(*
SPDX-FileCopyrightText: © 2026 Oleksandr Tiutyk <trofimich@gmail.com>
SPDX-License-Identifier: MIT
License: https://opensource.org/license/mit
*)

(*!
<summary>Mock leaf for lifecycle hooks, I/O phases, initialization/reset faults and event routing.</summary>
*)

FUNCTION_BLOCK MockLeafAutomationComponent EXTENDS TOF_Automation.InputOutputLeafAutomationComponent
VAR_INPUT
	//! <summary>Raises one output fault after the output call has been counted.</summary>
	ThrowOnNextOutput : BOOL;
	//! <summary>Raises one fault during input acquisition.</summary>
	ThrowOnNextInput : BOOL;
END_VAR
VAR_STAT
	{attribute 'hide'}
	_ClassName : STRING := __POUNAME();
END_VAR
VAR
	{attribute 'hide'}
	_InitializeCount : INT;
	{attribute 'hide'}
	_WorkingCount : INT;
	{attribute 'hide'}
	_ProcessInputCount : INT;
	{attribute 'hide'}
	_ProcessOutputCount : INT;
	{attribute 'hide'}
	_ResetCount : INT;
	{attribute 'hide'}
	_StopCount : INT;
	{attribute 'hide'}
	_EnableCount : INT;
	{attribute 'hide'}
	_DisableCount : INT;
	{attribute 'hide'}
	_EventReceivedCount : INT;
	{attribute 'hide'}
	_LastReceivedEventId : INT;
	{attribute 'hide'}
	_StopPropagationOnEvent : BOOL;
	{attribute 'hide'}
	_InitReturnValue : BOOL := TRUE;
	{attribute 'hide'}
	_FailOnWorking : BOOL;
	_ThrowOnInitializing : BOOL;
	_ThrowOnReset : BOOL;
	_RecoverCount : INT;
	_ThrowOnRecover : BOOL;
	_ThrowOnEnable : BOOL;
	_ThrowOnDisable : BOOL;
END_VAR

{attribute 'monitoring' := 'call'}
PROPERTY ClassName : REFERENCE TO STRING
GET
ClassName REF= _ClassName;
END_GET
END_PROPERTY

{attribute 'monitoring' := 'call'}
PROPERTY DisableCount : INT
GET
DisableCount := _DisableCount;
END_GET
END_PROPERTY

{attribute 'monitoring' := 'call'}
PROPERTY EnableCount : INT
GET
EnableCount := _EnableCount;
END_GET
END_PROPERTY

{attribute 'monitoring' := 'call'}
PROPERTY EventReceivedCount : INT
GET
EventReceivedCount := _EventReceivedCount;
END_GET
END_PROPERTY

{attribute 'monitoring' := 'call'}
PROPERTY FailOnWorking : BOOL
GET
FailOnWorking := _FailOnWorking;
END_GET
SET
_FailOnWorking := FailOnWorking;
END_SET
END_PROPERTY

METHOD FB_init : BOOL
VAR_INPUT
	bInitRetains : BOOL; // TRUE: the retain variables are initialized (reset warm / reset cold)
	bInCopyCode : BOOL;  // TRUE: the instance will be copied to the copy code afterward (online change)
	name : WSTRING;
	parent : TOF_Automation.IParentAutomationComponent;
END_VAR
END_METHOD

{attribute 'monitoring' := 'call'}
PROPERTY InitializeCount : INT
GET
InitializeCount := _InitializeCount;
END_GET
END_PROPERTY

{attribute 'monitoring' := 'call'}
PROPERTY InitReturnValue : BOOL
GET
InitReturnValue := _InitReturnValue;
END_GET
SET
_InitReturnValue := InitReturnValue;
END_SET
END_PROPERTY

{attribute 'monitoring' := 'call'}
PROPERTY LastReceivedEventId : INT
GET
LastReceivedEventId := _LastReceivedEventId;
END_GET
END_PROPERTY

{attribute 'monitoring' := 'call'}
PROPERTY NamespaceName : REFERENCE TO STRING
GET
NamespaceName REF= CurrentNamespace.Name;
END_GET
END_PROPERTY

(*!
<summary>Records the OnDisable call and optionally injects an exception.</summary>
*)
METHOD PROTECTED OnDisable
_DisableCount := _DisableCount + 1;

IF _ThrowOnDisable THEN
	TOF_Core.Exceptions.ThrowStandard(
		sourceNamespaceName := NamespaceName,
		sourceClassName := ClassName,
		sourcePOUName := __POUNAME(),
		sourcePosition := __POSITION(),
		message := "Injected OnDisable failure."
	);
END_IF
END_METHOD

(*!
<summary>Records the OnEnable call and optionally injects an exception.</summary>
*)
METHOD PROTECTED OnEnable
_EnableCount := _EnableCount + 1;

IF _ThrowOnEnable THEN
	TOF_Core.Exceptions.ThrowStandard(
		sourceNamespaceName := NamespaceName,
		sourceClassName := ClassName,
		sourcePOUName := __POUNAME(),
		sourcePosition := __POSITION(),
		message := "Injected OnEnable failure."
	);
END_IF
END_METHOD

METHOD OnEventReceived
VAR_INPUT
	event : TOF_Core.IEvent;
END_VAR
VAR_OUTPUT
	stopPropagation : BOOL;
END_VAR
VAR
	mockEv : POINTER TO MockAutomationEvent;
END_VAR
_EventReceivedCount := _EventReceivedCount + 1;

IF __QUERYPOINTER(event, mockEv) THEN
	_LastReceivedEventId := mockEv^.EventId;
END_IF

stopPropagation := _StopPropagationOnEvent;
END_METHOD

(*!
<summary>Records the OnInitializing call and optionally injects an exception.</summary>
<description>
The exception exercises production conversion into a copied component error; the hook does not own it.
</description>
*)
METHOD PROTECTED OnInitializing : BOOL
_InitializeCount := _InitializeCount + 1;

IF _ThrowOnInitializing THEN
	TOF_Core.Exceptions.ThrowStandard(
		sourceNamespaceName := NamespaceName,
		sourceClassName := ClassName,
		sourcePOUName := __POUNAME(),
		sourcePosition := __POSITION(),
		message := "Injected OnInitializing failure."
	);
END_IF

OnInitializing := _InitReturnValue;
END_METHOD

(*! <summary>Counts input calls and raises an armed input fault once.</summary> *)
METHOD PROTECTED OnProcessInput
_ProcessInputCount := _ProcessInputCount + 1;

IF ThrowOnNextInput THEN
	ThrowOnNextInput := FALSE;
	TOF_Core.Exceptions.ThrowStandard(
		sourceNamespaceName := NamespaceName,
		sourceClassName := ClassName,
		sourcePOUName := __POUNAME(),
		sourcePosition := __POSITION(),
		message := "Injected input failure"
	);
END_IF
END_METHOD

(*! <summary>Counts output calls and optionally injects a one-shot fault after the observed effect.</summary> *)
METHOD PROTECTED OnProcessOutput
_ProcessOutputCount := _ProcessOutputCount + 1;

IF ThrowOnNextOutput THEN
	ThrowOnNextOutput := FALSE;
	TOF_Core.Exceptions.ThrowStandard(
		sourceNamespaceName := NamespaceName,
		sourceClassName := ClassName,
		sourcePOUName := __POUNAME(),
		sourcePosition := __POSITION(),
		message := "Injected output failure"
	);
END_IF
END_METHOD

(*!
<summary>Records the OnRecover call and optionally injects an exception.</summary>
*)
METHOD PROTECTED OnRecover
_RecoverCount := _RecoverCount + 1;

IF _ThrowOnRecover THEN
	TOF_Core.Exceptions.ThrowStandard(
		sourceNamespaceName := NamespaceName,
		sourceClassName := ClassName,
		sourcePOUName := __POUNAME(),
		sourcePosition := __POSITION(),
		message := "Injected OnRecover failure."
	);
END_IF
END_METHOD

(*!
<summary>Records the OnReset call and optionally injects an exception.</summary>
<description>
The exception exercises production conversion into a copied component error; the hook does not own it.
</description>
*)
METHOD PROTECTED OnReset
_ResetCount := _ResetCount + 1;

IF _ThrowOnReset THEN
	TOF_Core.Exceptions.ThrowStandard(
		sourceNamespaceName := NamespaceName,
		sourceClassName := ClassName,
		sourcePOUName := __POUNAME(),
		sourcePosition := __POSITION(),
		message := "Injected OnReset failure."
	);
END_IF
END_METHOD

METHOD PROTECTED OnStopped
_StopCount := _StopCount + 1;
END_METHOD

METHOD PROTECTED OnWorking
_WorkingCount := _WorkingCount + 1;

IF _FailOnWorking THEN
	TOF_Core.Exceptions.ThrowStandard(
		sourceNamespaceName := NamespaceName,
		sourceClassName := ClassName,
		sourcePOUName := __POUNAME(),
		sourcePosition := __POSITION(),
		message := "Mock leaf failure on working"
	);
END_IF
END_METHOD

{attribute 'monitoring' := 'call'}
PROPERTY ProcessInputCount : INT
GET
ProcessInputCount := _ProcessInputCount;
END_GET
END_PROPERTY

{attribute 'monitoring' := 'call'}
PROPERTY ProcessOutputCount : INT
GET
ProcessOutputCount := _ProcessOutputCount;
END_GET
END_PROPERTY

{attribute 'monitoring' := 'call'}
PROPERTY ResetCount : INT
GET
ResetCount := _ResetCount;
END_GET
END_PROPERTY

{attribute 'monitoring' := 'call'}
PROPERTY SelfSize : ULINT
GET
SelfSize := XSIZEOF(THIS^);
END_GET
END_PROPERTY

{attribute 'monitoring' := 'call'}
PROPERTY StopCount : INT
GET
StopCount := _StopCount;
END_GET
END_PROPERTY

{attribute 'monitoring' := 'call'}
PROPERTY StopPropagationOnEvent : BOOL
GET
StopPropagationOnEvent := _StopPropagationOnEvent;
END_GET
SET
_StopPropagationOnEvent := StopPropagationOnEvent;
END_SET
END_PROPERTY

{attribute 'monitoring' := 'call'}
PROPERTY WorkingCount : INT
GET
WorkingCount := _WorkingCount;
END_GET
END_PROPERTY

(*!
<summary>Controls the initialization-hook failure injected by regression tests.</summary>
*)
{attribute 'monitoring' := 'call'}
PROPERTY ThrowOnInitializing : BOOL
GET
ThrowOnInitializing := _ThrowOnInitializing;
END_GET
SET
_ThrowOnInitializing := ThrowOnInitializing;
END_SET
END_PROPERTY

(*!
<summary>Controls the reset-hook failure injected by regression tests.</summary>
*)
{attribute 'monitoring' := 'call'}
PROPERTY ThrowOnReset : BOOL
GET
ThrowOnReset := _ThrowOnReset;
END_GET
SET
_ThrowOnReset := ThrowOnReset;
END_SET
END_PROPERTY

(*!
<summary>Gets the number of OnRecover calls recorded by this mock leaf.</summary>
*)
{attribute 'monitoring' := 'call'}
PROPERTY RecoverCount : INT
GET
RecoverCount := _RecoverCount;
END_GET
END_PROPERTY

(*!
<summary>Controls the disable-hook failure injected by regression tests.</summary>
*)
{attribute 'monitoring' := 'call'}
PROPERTY ThrowOnDisable : BOOL
GET
ThrowOnDisable := _ThrowOnDisable;
END_GET
SET
_ThrowOnDisable := ThrowOnDisable;
END_SET
END_PROPERTY

(*!
<summary>Controls the enable-hook failure injected by regression tests.</summary>
*)
{attribute 'monitoring' := 'call'}
PROPERTY ThrowOnEnable : BOOL
GET
ThrowOnEnable := _ThrowOnEnable;
END_GET
SET
_ThrowOnEnable := ThrowOnEnable;
END_SET
END_PROPERTY

(*!
<summary>Controls the recover-hook failure injected by regression tests.</summary>
*)
{attribute 'monitoring' := 'call'}
PROPERTY ThrowOnRecover : BOOL
GET
ThrowOnRecover := _ThrowOnRecover;
END_GET
SET
_ThrowOnRecover := ThrowOnRecover;
END_SET
END_PROPERTY

(*!
<summary>Exercises the inherited exception handler with a borrowed diagnostic in the fixture's current state.</summary>
<param name="exception">Task-local exception that remains live for the call.</param>
<param name="reaction">Runtime reaction to apply.</param>
*)
METHOD ApplyExceptionReaction
VAR_INPUT
	exception : TOF_Core.IException;
	reaction : TOF_Core.EXCEPTION_REACTION;
END_VAR
ProcessException(exception := exception, exceptionReaction := reaction, exceptionSourceHint := "Injected primary failure");
END_METHOD

END_FUNCTION_BLOCK

(* stored: Version 1.1.0.1, ProductVersion 3.1.4026.21
   POU MockLeafAutomationComponent: Id {9b7b3daa-f346-4584-a906-6da16219c11f}, SpecialFunc None
   Folder Methods to override: Id {612da229-f7d8-494f-8591-082c05072b3f}
   Folder Properties for tests: Id {ccac3e62-bc35-4f89-a40e-c876ffb73e34}
   Property ClassName: Id {d5c4d5ee-cde5-4df4-8cbd-46cced7d5454}
   Get Get: Id {5415ed35-e09f-4119-8198-c8575e6b1ab5}
   Property DisableCount: Id {bbaaaf6d-9d95-455d-b78d-b03325aec8ca}
   Get Get: Id {16fe8a7f-cfad-4055-9144-48f18add74a5}
   Property EnableCount: Id {8454a8af-ef78-4131-b582-201baa06e86e}
   Get Get: Id {489c43e4-5062-4c21-8691-e46ab060d4b5}
   Property EventReceivedCount: Id {803a68c5-6fea-4132-9ec0-3eab19c89d39}
   Get Get: Id {bd615afb-6d2f-41d6-88ec-30cdcef21a93}
   Property FailOnWorking: Id {4ac1dd38-5fe7-40fa-b603-9534ebe240bd}
   Get Get: Id {da42525c-79be-4472-94c1-fd35af010373}
   Set Set: Id {a2eba756-0bc3-4394-adfb-aa16c4171792}
   Method FB_init: Id {2ce54561-f6b4-4f38-b28c-e9e2d5ba5306}
   Property InitializeCount: Id {ff7ba116-c221-4cd9-9799-5b16792aeb45}
   Get Get: Id {018cb720-e3f7-4649-8b67-bed593899c5b}
   Property InitReturnValue: Id {69a85714-ee34-4f3d-80b7-d8d28b5786a9}
   Get Get: Id {c7fd5de5-7d8a-4d20-b545-b2cc79f89fe3}
   Set Set: Id {b19d322b-4ce8-4aa2-a823-6e081aa50e60}
   Property LastReceivedEventId: Id {b620503e-4868-4d7f-8ccf-6c554061f9ae}
   Get Get: Id {d7856263-a660-4787-a01c-8114042f908c}
   Property NamespaceName: Id {56d74b1c-f6c9-459f-9c64-e87f22404f29}
   Get Get: Id {8d20768a-1d4c-48d9-b2ea-aa35fdbec9c1}
   Method OnDisable: Id {d2427892-1a02-494e-bfe1-cdea7c7139be}
   Method OnEnable: Id {536c9e62-ae74-4c2a-be87-73caf5b19d2b}
   Method OnEventReceived: Id {0c87de76-5092-4e69-b2f2-bf3d5f3a3ac8}
   Method OnInitializing: Id {6fb51265-efad-48f5-a686-62ad9bd26b0a}
   Method OnProcessInput: Id {16a990da-11aa-4e60-bc1c-debaa2275464}
   Method OnProcessOutput: Id {13d5c65e-afd4-4d9c-a902-9000ddab6569}
   Method OnRecover: Id {20ebc6f7-f14d-42b0-bb2d-a84122dbeec8}
   Method OnReset: Id {1a42e8fd-4f72-4198-b9e9-5592070c737e}
   Method OnStopped: Id {b3148cc2-962a-490b-ba15-a96998f300aa}
   Method OnWorking: Id {739d0f66-08d3-465b-b7a1-458c0649f3ae}
   Property ProcessInputCount: Id {cbed7228-ef36-4fe8-afdf-425804d6c226}
   Get Get: Id {8b0f41f9-c2a4-4146-a82d-aba8bbf96cdb}
   Property ProcessOutputCount: Id {21ae72e0-b5af-4c1d-a75e-712952e8ecde}
   Get Get: Id {5f5940e0-d2b8-4a63-86b7-32565b7d7bf5}
   Property ResetCount: Id {dd549592-888a-4fd2-a904-1aa49b5cf483}
   Get Get: Id {5f28075a-c278-40f9-8ebc-71090e887d37}
   Property SelfSize: Id {623558a3-feec-4048-83fd-7afec0f97f19}
   Get Get: Id {d5d338c0-7d96-4e75-ae51-a5b4c7ddb7c2}
   Property StopCount: Id {6f90d479-70eb-43dd-a7d6-4c9abf5b97b4}
   Get Get: Id {10542a9e-26f1-47e9-ad6e-714891b57965}
   Property StopPropagationOnEvent: Id {0368d1d6-d4ba-4ae7-95d4-c46fb1019742}
   Get Get: Id {2d37d725-4fe9-48d6-8aa0-963c2d1a5188}
   Set Set: Id {17c8c87e-07cd-49ed-a163-45a2585fc087}
   Property WorkingCount: Id {acd0aabc-538a-45c9-8870-7bb40400c830}
   Get Get: Id {25c6fb63-a350-4fe0-9ada-f16c40e49355}
   Property ThrowOnInitializing: Id {112053f4-0cbc-41b5-a06a-87a87a46364f}
   Get Get: Id {ffe3d562-5540-4e3e-ad76-d837a6dde8a4}
   Set Set: Id {c1a76dd8-0de4-44b5-89f1-eea061a87c48}
   Property ThrowOnReset: Id {9ea1bff4-c2c6-46f6-b244-a52eb26b2f46}
   Get Get: Id {91d419db-0fd3-4005-a532-2471f9189792}
   Set Set: Id {841ec3fb-3c6d-42ce-bc1d-07c4611e638f}
   Property RecoverCount: Id {bc1a696f-03e8-4bf2-811e-8633f58a1f71}
   Get Get: Id {707352ed-757e-4840-9178-5cf678c3cc50}
   Property ThrowOnDisable: Id {5667a825-c8c5-4181-9533-c2e45376dcc4}
   Get Get: Id {5b90252b-5e02-4bce-a79a-b51fd2188211}
   Set Set: Id {caef36ea-6e29-461b-91d9-a1e08aa4597c}
   Property ThrowOnEnable: Id {f0937ab9-60ab-42c2-a656-6ea7e8028419}
   Get Get: Id {7568e807-85f4-4924-a05c-884344dc070f}
   Set Set: Id {b316f523-9150-440a-a5aa-3a7cfce64e92}
   Property ThrowOnRecover: Id {5b8e6502-ae6e-44bb-95fa-7aa83026891b}
   Get Get: Id {9ae2ed04-50a6-4915-aed1-7525fac24f43}
   Set Set: Id {7b5fc291-25e6-46f7-ba3d-7074f72ad46b}
   Method ApplyExceptionReaction: Id {5c891c44-9149-4457-adb2-6048d59c3797} *)
